(* IEC 61131-3 sources: SRCI_CLIENT_PLC/RobotLibrary/Library/POUs/_internal, 1 file *)

(* ---- ActiveCommandRegisterFB.st ---- *)
FUNCTION_BLOCK ActiveCommandRegisterFB EXTENDS RobotLibraryLogFB
// -------------------------------------------------------------------------
//  SRCI Robot Library
// -------------------------------------------------------------------------
//
//  Object:      ActiveCommandRegisterFB
//  Author:      Thorsten Brach
//  Date:        2024-06-01
//
//  Description:
//
//
//  Copyright:
//    (C) 2024 Thorsten Brach. All rights reserved
//             Licensed under the MIT License.
//
//  Disclaimer:
//    This project is provided without any guarantee and can be used for
//    private and commercial purposes. Any use is at the user’s
//    own risk and responsibility.
//
// -------------------------------------------------------------------------
VAR_INPUT
  /// Active Command Register
  Register            : ARRAY [1..RobotLibraryParameter.ACTIVE_CMD_REGISTER_ENTRIES_MAX] OF AxesGroupAcyclicAcrEntry;
  /// System Time
  SystemTime          : SystemTime;
  /// usable size of the arc register
  RegisterSize        : DINT := RobotLibraryParameter.ACTIVE_CMD_REGISTER_ENTRIES_MAX;
END_VAR

VAR_OUTPUT
  /// Execution Order List
  ExecutionOrderList    : ARRAY [1..RobotLibraryParameter.ACTIVE_CMD_REGISTER_ENTRIES_MAX] OF DINT;
  /// Current amount of used registers
  CurrentAcrUsageCount  : DINT;
  /// Current percent of used registers
  CurrentAcrUsagePercent : REAL;
END_VAR

VAR
  /// temporarty Active Command Register
  TmpRegister                 : ARRAY [1..RobotLibraryParameter.ACTIVE_CMD_REGISTER_ENTRIES_MAX] OF AxesGroupAcyclicAcrEntry;
  /// last used unique ID
  LastUniqueID                : UINT;
  /// Warning for ACR usage at 80%
  WarningAcrUsage             : R_TRIG;
END_VAR

VAR CONSTANT
  /// Active command
  ACTIVE_CMD           : UDINT := 1;
  /// Buffered command
  BUFFER_CMD           : UDINT := 2;
  /// Empty ACR entry
  EMPTY_ACR_ENTRY      : AxesGroupAcyclicAcrEntry := (State := ActiveCommandRegisterState.IS_FREE);
  /// Empty command entry
  EMPTY_CMD_ENTRY      : AxesGroupAcyclicAcrEntryCmdBuffer := (State := BufferStateCmd.EMPTY);
  /// constant for byte index of priority in payload
  PRIORITY_IDX         : BYTE := 3;
  /// bitmask to mask the priority out of the halfbyte
  PRIORITY_BIT_MASK    : BYTE := 2#000_1111;
END_VAR

  ManageRegister();

  UpdateExecutionOrderList();

END_FUNCTION_BLOCK

METHOD PUBLIC AddCmd : UDINT
VAR_INPUT
  /// Pointer to the corresponding command-FB to enable a callback mechanism
  pCommandFB        : POINTER TO RobotLibraryBaseFB;
END_VAR

VAR
  /// internal index for loops
 _regIdx            : DINT;
  /// internal command type
 _cmdType           : CmdType;
  /// log message
 _messageLog        : AlarmMessage;
  /// flag for free register found
 _freeRegisterFound : BOOL;
  /// internal Acr error
 _errorAcrEntry     : WORD := RobotLibraryErrorIdEnum.ERR_NO_FREE_ACR_ENTRY;
END_VAR

  // ST-FIX F48: a command with a parameter error of the block is not added
  IF ( pCommandFB <> 0 )
  THEN
    IF (( pCommandFB^.ErrorID = RobotLibraryErrorIdEnum.ERR_INVALID_PARAM_EXECUTION_MODE ) OR
        ( pCommandFB^.ErrorID = RobotLibraryErrorIdEnum.ERR_PROCESSINGMODE_NOT_DEFINED   ))
    THEN
      AddCmd := 0;
      RETURN;
    END_IF
  END_IF

  // calculate the used length of the ACR
  FOR _regIdx := 1 TO RegisterSize
  DO
    IF ( Register[_regIdx].State = ActiveCommandRegisterState.IS_FREE )
    THEN
      Register[_regIdx].State      := ActiveCommandRegisterState.IS_PROCESSING;
      Register[_regIdx].UniqueID   := DINT_TO_UINT(_regIdx);
      Register[_regIdx].pCommandFB := pCommandFB;

      // check pointer to command FB
      IF ( Register[_regIdx].pCommandFB <> RobotLibraryConstants.NULL_POINTER )
      THEN
        Register[_regIdx].Command[RobotLibraryConstants.ACTIVE_CMD].Timestamp  := SystemTime;

        Register[_regIdx].Command[RobotLibraryConstants.ACTIVE_CMD].Payload    := pCommandFB^.CommandData.Payload;
        Register[_regIdx].Command[RobotLibraryConstants.ACTIVE_CMD].PayloadLen := pCommandFB^.CommandData.PayloadLen;
        Register[_regIdx].Command[RobotLibraryConstants.ACTIVE_CMD].PayLoadPtr := 0;
        Register[_regIdx].Command[RobotLibraryConstants.ACTIVE_CMD].State      := BufferStateCmd.CREATED;
      END_IF

      // set flag for free register found
     _freeRegisterFound := TRUE;

      // Increment Current used register counter
      CurrentAcrUsageCount := CurrentAcrUsageCount + 1;

      // return Unique ID
      AddCmd := Register[_regIdx].UniqueID;

      // Get CmdType from payload
      SysDepMemCpy( pDest := ADR(_cmdType), pSrc := ADR(pCommandFB^.CommandData.Payload), DataLen := SIZEOF(_cmdType));

      // Create log entry
      CreateLogMessagePara2 ( Timestamp   := SystemTime,
                              MessageType := MessageType.CMD,
                              Severity    := Severity.INFO,
                              MessageCode := 0,
                              MessageText := 'ACR-ID [{1}]: Added  Command-Payload of CmdType <{2}>',
                              Para1       :=  DINT_TO_STRING(_regIdx),
                              Para2       :=  CMD_TYPE_TO_STRING(SwapUint(_cmdType)));
      EXIT;
    END_IF
  END_FOR

  // Check a free register could be found ?
  IF ( NOT _freeRegisterFound )
  THEN
    // set error in Command FB
    IF ( pCommandFB <> RobotLibraryConstants.NULL_POINTER )
    THEN
      SysDepMemCpy( pDest   := ADR   ( pCommandFB^.ErrorID ),
                    pSrc    := ADR   ( _errorAcrEntry      ),
                    DataLen := SIZEOF( _errorAcrEntry      ));
    END_IF

    // Create log entry
    CreateLogMessagePara1 ( Timestamp   := SystemTime,
                            MessageType := MessageType.CMD,
                            Severity    := Severity.FATAL_ERROR,
                            MessageCode := 0,
                            MessageText := 'Not possible to add CMD <{1}> to ACR - NO FREE REGISTER FOUND ! -> STOPPING SRCI INTERFACE...',
                            Para1       :=  CMD_TYPE_TO_STRING(SwapUint(_cmdType)));
  END_IF

END_METHOD

METHOD AddRsp : UDINT
VAR_INPUT
  /// Response
  Rsp : TelegramRobToPlcFragment;
END_VAR
VAR
  /// internal index for loops
 _Idx             : DINT;
  /// internal registen index
 _regIdx          : DINT;
  /// internal command type
 _cmdType         : CmdType;
  /// internal FragmentAction
 _fragmentAction  :  FragmentAction;
  /// internal command message state
 _cmdMessageState : CmdMessageState;
  /// internal flag for CmdID found
 _found           : BOOL;
END_VAR

  FOR _regIdx := 1 TO RegisterSize
  DO
    IF ( Register[_regIdx].UniqueID = Rsp.Header.CmdID )
    THEN
      // CmdID was found in the ACR
     _found := TRUE;
      // convert to fragment action
     _fragmentAction := ByteToFragmentAction(Rsp.Header.FragmentAction);

      // delete response
      IF ( _fragmentAction.Clear )
      THEN
        SysDepMemSet( pDest := ADR(Register[_regIdx].Response[ACTIVE_CMD]), Value := 0, DataLen := SIZEOF(Register[_regIdx].Response[ACTIVE_CMD]));
      END_IF

      // add payload to response
      FOR _idx := Rsp.Header.PayloadPointer TO  Rsp.Header.PayloadPointer + Rsp.Header.PayloadLength -1
      DO
        Register[_regIdx].Response[ACTIVE_CMD].Timestamp     := SystemTime;
        Register[_regIdx].Response[ACTIVE_CMD].State         := BufferStateRsp.RECEIVING;
        Register[_regIdx].Response[ACTIVE_CMD].PayloadLen    := Register[_regIdx].Response[ACTIVE_CMD].PayloadLen + 1;
        Register[_regIdx].Response[ACTIVE_CMD].Payload[_idx] := Rsp.Command.Payload[_idx];
      END_FOR

      // Get current message state
     _cmdMessageState := GetHalfeByteLo    (Value  := Register[_regIdx].Response[ACTIVE_CMD].Payload[0]);
      // Get command type from payload
     _cmdType         := CombineBytesToUint(HiByte := Register[_regIdx].Command [ACTIVE_CMD].Payload[0],
                                            LoByte := Register[_regIdx].Command [ACTIVE_CMD].Payload[1]);

      // Create log entry
      CreateLogMessagePara3 ( Timestamp   := SystemTime,
                              MessageType := MessageType.CMD,
                              Severity    := Severity.INFO,
                              MessageCode := 0,
                              MessageText := 'ACR-ID [{1}]: Added Response-Payload of CmdType <{2}> with State = {3}',
                              Para1       :=  DINT_TO_STRING(_regIdx),
                              Para2       :=  CMD_TYPE_TO_STRING(_cmdType),
                              Para3       :=  CMD_MESSAGE_STATE_TO_STRING(_cmdMessageState));

      IF ( _fragmentAction.Complete )
      THEN
        // set response state
        Register[_regIdx].Response[ACTIVE_CMD].State := BufferStateRsp.RECEIVED;

        // Check current message state and tag the register state as IS_FINAL, if needed
        IF ( _cmdMessageState >= CmdMessageState.DONE)
        THEN
          Register[_regIdx].State := ActiveCommandRegisterState.IS_FINAL;

          // get command type from payload
         _cmdType := CombineBytesToUint(HiByte := Register[_regIdx].Command[ACTIVE_CMD].Payload[0],
                                        LoByte := Register[_regIdx].Command[ACTIVE_CMD].Payload[1]);

          // Create log entry
          CreateLogMessagePara3( Timestamp   := SystemTime,
                                 MessageType := MessageType.CMD,
                                 Severity    := Severity.INFO,
                                 MessageCode := 0,
                                 MessageText := 'ACR-ID [{1}]: Detected Response-Payload of CmdType <{2}> has reached final state <{3}>',
                                 Para1       :=  DINT_TO_STRING(_regIdx),
                                 Para2       :=  CMD_TYPE_TO_STRING(_cmdType),
                                 Para3       :=  CMD_MESSAGE_STATE_TO_STRING(_cmdMessageState));

          // Exit the loop
        END_IF
      END_IF

      // Check Response received complete ?
      IF ( Register[_regIdx].Response[ACTIVE_CMD].State = BufferStateRsp.RECEIVED)
      THEN
        // update state
        Register[_regIdx].Response[ACTIVE_CMD].State := BufferStateRsp.PROCESSED;
        // callback CommandFB
        Register[_regIdx].pCommandFB^.CallBack(RspData := Register[_regIdx].Response[ACTIVE_CMD],TimeStamp := SystemTime);
      END_IF

      EXIT;
    END_IF
  END_FOR

  // Check CmdID was found in the ACR ?
  IF ( NOT _found )
  THEN
    // Create log entry
    CreateLogMessagePara2 ( Timestamp   := SystemTime,
                            MessageType := MessageType.CMD,
                            Severity    := Severity.WARNING,
                            MessageCode := 0,
                            MessageText := 'ACR-ID [?]: Response-Payload of CmdID <{1}> with State = {2} received, but no matching ACR entry found',
                            Para1       :=  UINT_TO_STRING(Rsp.Header.CmdID),
                            Para2       :=  CMD_MESSAGE_STATE_TO_STRING(_cmdMessageState));
  END_IF

END_METHOD

METHOD FB_init : BOOL
VAR_INPUT
  bInitRetains : BOOL; // if TRUE, the retain variables are initialized (warm start / cold start)
  bInCopyCode : BOOL;  // if TRUE, the instance afterwards gets moved into the copy code (online change)
END_VAR

  MyType := 'ActiveCommandRegisterFB';

END_METHOD

METHOD PRIVATE ManageRegister
VAR
  /// internal index
 _regIdx          : DINT;
  /// internal command type
 _cmdType         : CmdType;
  /// internal command message state
 _cmdMessageState : CmdMessageState;
END_VAR

  FOR _regIdx := 1 TO RegisterSize
  DO
    // Check pointer to command FB is valid ?
    IF ( Register[_regIdx].pCommandFB <> RobotLibraryConstants.NULL_POINTER)
    THEN

      // Check apply Cmd parameter update ?
      IF (( Register[_regIdx].Command[ACTIVE_CMD].State = BufferStateCmd.PROCESSED        ) AND
          ( Register[_regIdx].Command[BUFFER_CMD].State = BufferStateCmd.UPDATE_AVAILABLE ))
      THEN
        Register[_regIdx].Command[ACTIVE_CMD] := Register[_regIdx].Command[BUFFER_CMD];
        Register[_regIdx].Command[BUFFER_CMD] := EMPTY_CMD_ENTRY;

        // get command type from payload
       _cmdType := CombineBytesToUint(HiByte := Register[_regIdx].Command[ACTIVE_CMD].Payload[0],
                                      LoByte := Register[_regIdx].Command[ACTIVE_CMD].Payload[1]);

        // Create log entry
        CreateLogMessagePara2 ( Timestamp   := SystemTime,
                                MessageType := MessageType.CMD,
                                Severity    := Severity.INFO,
                                MessageCode := 0,
                                MessageText := 'ACR-ID [{1}]: Moved BUFFER_CMD to ACTIVE_CMD, CmdType <{2}>',
                                Para1       :=  DINT_TO_STRING(_regIdx),
                                Para2       :=  CMD_TYPE_TO_STRING(_cmdType));

      END_IF

      (*
      // Check Response received ?
      IF ( Register[_regIdx].Response[ACTIVE_CMD].State = BufferStateRsp.RECEIVED)
      THEN
        // update state
        Register[_regIdx].Response[ACTIVE_CMD].State := BufferStateRsp.PROCESSED;
        // callback CommandFB
        Register[_regIdx].pCommandFB^.CallBack(RspData := Register[_regIdx].Response[ACTIVE_CMD],TimeStamp := SystemTime);
      END_IF
      *)

      // delete entries with State.IS_Final
      IF ( Register[_regIdx].State = ActiveCommandRegisterState.IS_FINAL )
      THEN
        // get command type from payload
       _cmdType := CombineBytesToUint(HiByte := Register[_regIdx].Command[ACTIVE_CMD].Payload[0],
                                      LoByte := Register[_regIdx].Command[ACTIVE_CMD].Payload[1]);

        // Get current message state
       _cmdMessageState := GetHalfeByteLo(Value := Register[_regIdx].Response[ACTIVE_CMD].Payload[0]);

        // Create log entry
        CreateLogMessagePara3( Timestamp   := SystemTime,
                               MessageType := MessageType.CMD,
                               Severity    := Severity.INFO,
                               MessageCode := 0,
                               MessageText := 'ACR-ID [{1}]: Deleted ACR-Entry of CmdType <{2}> with State = {3}, because of Final-State was reached',
                               Para1       :=  DINT_TO_STRING(_regIdx),
                               Para2       :=  CMD_TYPE_TO_STRING(_cmdType),
                               Para3       :=  CMD_MESSAGE_STATE_TO_STRING(_cmdMessageState));

        // delete register entry
        Register[_regIdx] := EMPTY_ACR_ENTRY;

        // decrement current used register counter
        CurrentAcrUsageCount := CurrentAcrUsageCount - 1;
      END_IF
    END_IF
  END_FOR

  // Calculate percent of register usage
  IF ( CurrentAcrUsageCount > 0)
  THEN
    CurrentAcrUsagePercent :=  (DINT_TO_REAL(CurrentAcrUsageCount) / DINT_TO_REAL(RegisterSize)) * 100.0;
  ELSE
    CurrentAcrUsagePercent := 0.0;
  END_IF

  // build rising edge for arc usage over 80%
  WarningAcrUsage( CLK := CurrentAcrUsagePercent > RobotLibraryParameter.ACR_USAGE_WARNING_LIMIT );

  IF ( WarningAcrUsage.Q )
  THEN
    // Create log entry
    CreateLogMessagePara4( Timestamp   := SystemTime,
                           MessageType := MessageType.CMD,
                           Severity    := Severity.WARNING,
                           MessageCode := 0,
                           MessageText := 'ACR Register usage has reached the warning limit ({1}): {2}/{3} = {4}%',
                           Para1       :=  REAL_TO_STRING(RobotLibraryParameter.ACR_USAGE_WARNING_LIMIT),
                           Para2       :=  DINT_TO_STRING(CurrentAcrUsageCount),
                           Para3       :=  DINT_TO_STRING(RegisterSize),
                           Para4       :=  REAL_TO_STRING(CurrentAcrUsagePercent));
  END_IF

END_METHOD

PROPERTY PUBLIC NotifyParameterChanged : UDINT

SET
VAR
  /// internal register index
 _regIdx  : DINT;
  /// internal command type
 _cmdType : CmdType;
END_VAR

  FOR _regIdx := 1 TO RobotLibraryParameter.ACTIVE_CMD_REGISTER_ENTRIES_MAX
  DO
    // check unique ID found ?
    IF ( Register[_regIdx].UniqueID = NotifyParameterChanged )
    THEN
      // ST-FIX F114: a parameter change before the command is sent (state CREATED) must not turn the new
      // command into a parameter update (it was never sent): the command keeps the parameters of the rising edge
      IF ( Register[_regIdx].Command[ACTIVE_CMD].State = BufferStateCmd.CREATED )
      THEN
        // Create log entry
        CreateLogMessagePara1 ( Timestamp   := SystemTime,
                                MessageType := MessageType.CMD,
                                Severity    := Severity.INFO,
                                MessageCode := 0,
                                MessageText := 'ACR-ID [{1}]: Cmd-Parameter changed before the command was sent -> ignored',
                                Para1       :=  DINT_TO_STRING(_regIdx));
      ELSIF (( Register[_regIdx].Command[ACTIVE_CMD].State <> BufferStateCmd.SENDING   ) AND
             ( Register[_regIdx].Command[ACTIVE_CMD].State <> BufferStateCmd.PROCESSED ))
      THEN
        // Check pointer is valid ?
        IF ( Register[_regIdx].pCommandFB <> RobotLibraryConstants.NULL_POINTER )
        THEN
          // add to send register
          Register[_regIdx].Command[ACTIVE_CMD].Timestamp  := SystemTime;
          Register[_regIdx].Command[ACTIVE_CMD].State      := BufferStateCmd.UPDATE_AVAILABLE;
          Register[_regIdx].Command[ACTIVE_CMD].Payload    := Register[_regIdx].pCommandFB^.CommandData.Payload;
          Register[_regIdx].Command[ACTIVE_CMD].PayloadLen := Register[_regIdx].pCommandFB^.CommandData.PayloadLen;

          // get command type from payload
         _cmdType := CombineBytesToUint(HiByte := Register[_regIdx].pCommandFB^.CommandData.Payload[0],
                                        LoByte := Register[_regIdx].pCommandFB^.CommandData.Payload[1]);

          // Create log entry
          CreateLogMessagePara2 ( Timestamp   := SystemTime,
                                  MessageType := MessageType.CMD,
                                  Severity    := Severity.INFO,
                                  MessageCode := 0,
                                  MessageText := 'ACR-ID [{1}]: Updated Cmd-Parameter of CmdType <{2}> -> written to ACTIVE_CMD Index',
                                  Para1       :=  DINT_TO_STRING(_regIdx),
                                  Para2       :=  CMD_TYPE_TO_STRING(_cmdType));
        END_IF
      ELSE
        // Check pointer is valid ?
        IF ( Register[_regIdx].pCommandFB <> RobotLibraryConstants.NULL_POINTER )
        THEN
          // add to buffer register
          Register[_regIdx].Command[BUFFER_CMD].Timestamp  := SystemTime;
          Register[_regIdx].Command[BUFFER_CMD].State      := BufferStateCmd.UPDATE_AVAILABLE;
          Register[_regIdx].Command[BUFFER_CMD].Payload    := Register[_regIdx].pCommandFB^.CommandData.Payload;
          Register[_regIdx].Command[BUFFER_CMD].PayloadLen := Register[_regIdx].pCommandFB^.CommandData.PayloadLen;

          // get command type from payload
         _cmdType := CombineBytesToUint(HiByte := Register[_regIdx].pCommandFB^.CommandData.Payload[0],
                                        LoByte := Register[_regIdx].pCommandFB^.CommandData.Payload[1]);

          // Create log entry
          CreateLogMessagePara2 ( Timestamp   := SystemTime,
                                  MessageType := MessageType.CMD,
                                  Severity    := Severity.INFO,
                                  MessageCode := 0,
                                  MessageText := 'ACR-ID [{1}]: Updated Cmd-Parameter of CmdType <{2}> -> written to BUFFER_CMD Index',
                                  Para1       :=  DINT_TO_STRING(_regIdx),
                                  Para2       :=  CMD_TYPE_TO_STRING(_cmdType));
        END_IF
      END_IF

    END_IF
  END_FOR

END_SET

METHOD PUBLIC OnOnlineChange : DINT
VAR_INPUT
  /// unique ID
  UniqueID     : UDINT;
  /// Pointer to the corresponding command-FB to enable a callback mechanism
  pCommandFB   : POINTER TO RobotLibraryBaseFB;
END_VAR

VAR
  /// internal index for loops
 _regIdx : DINT;
END_VAR

  OnOnlineChange := -1;

  // Check command FB pointer is valid ?
  IF ( pCommandFB <> RobotLibraryConstants.NULL_POINTER)
  THEN
    FOR _regIdx := 1 TO RegisterSize
    DO
      // check unique ID found ?
      IF ( Register[_regIdx].UniqueID = UniqueID )
      THEN
        // update pointer to command FB
        Register[_regIdx].pCommandFB := pCommandFB;
        // Return result OK
        OnOnlineChange := RobotLibraryConstants.OK;
        EXIT;
      END_IF
    END_FOR
  END_IF

END_METHOD

METHOD PUBLIC RemoveCmd : DINT
VAR_INPUT
 /// unique ID
 UniqueID : UDINT;
END_VAR

VAR
  /// internal index
 _regIdx : DINT;
  /// internal command type
 _cmdType : CmdType;
END_VAR

  RemoveCmd := RobotLibraryConstants.HAS_ERROR;

  IF (UniqueID = 0)
  THEN
    UniqueID := UniqueID;
  END_IF

  FOR _regIdx := 1 TO RegisterSize
  DO
    // check unique ID found and not yet sended ?
    IF (( Register[_regIdx].UniqueID                  = UniqueID                        ) AND
        ( Register[_regIdx].Command[ACTIVE_CMD].State < BufferStateCmd.UPDATE_AVAILABLE ))
    THEN
      // Get CmdType from payload
      SysDepMemCpy( pDest := ADR(_cmdType), pSrc := ADR(Register[_regIdx].Command[ACTIVE_CMD].Payload), DataLen := SIZEOF(_cmdType));
      // delete register entry
      SysDepMemSet(pDest := ADR(Register[_regIdx]), Value := 0 , DataLen := SIZEOF(Register[_regIdx]));
      // decrement current used register counter
      CurrentAcrUsageCount := CurrentAcrUsageCount - 1;
      // Command successfull removed
      RemoveCmd := RobotLibraryConstants.OK;

      // Create log entry
      CreateLogMessagePara2 (  Timestamp   := SystemTime,
                               MessageType := MessageType.CMD,
                               Severity    := Severity.INFO,
                               MessageCode := 0,
                               MessageText := 'ACR-ID [{1}]: Removed CmdType <{2}>',
                               Para1       :=  DINT_TO_STRING(_regIdx),
                               Para2       :=  CMD_TYPE_TO_STRING(SwapUint(_cmdType)));
      EXIT;
    END_IF
  END_FOR

END_METHOD

METHOD PUBLIC Reset

  SysDepMemSet( ADR(Register), 0, SIZEOF(Register));

  CurrentAcrUsageCount   := 0;
  CurrentAcrUsagePercent := 0.0;

  // Create log entry
  CreateLogMessagePara1 ( Timestamp   := SystemTime,
                          MessageType := MessageType.CMD,
                          Severity    := Severity.INFO,
                          MessageCode := 0,
                          MessageText := 'ACR Registers has been reset and all entries deleted by Reset method call',
                          Para1       :=  '');

END_METHOD

METHOD PRIVATE UpdateExecutionOrderList
VAR
  /// temporary Active Command Register entry
  TmpRegisterEntry : AxesGroupAcyclicAcrEntry;
  /// temporary index
  TmpIndex         : DINT;
  /// internal index
  i                : DINT;
  /// internal index
  j                : DINT;
END_VAR

  // Reset temporary register
  SysDepMemSet(pDest := ADR(TmpRegister)       , Value := 0, DataLen := SIZEOF(TmpRegister));
  // Reset Execution Order List
  SysDepMemSet(pDest := ADR(ExecutionOrderList), Value := 0, DataLen := SIZEOF(ExecutionOrderList));
  // pre-set temporary register index
  j := 1;

  FOR i := 1 TO RegisterSize
  DO
    // add only entries which are not in status free and where datas must be processed
    IF (( Register[i].State                      > ActiveCommandRegisterState.IS_FREE ) AND
        ( Register[i].Command[ACTIVE_CMD].State <> BufferStateCmd.EMPTY               ) AND
        ( Register[i].Command[ACTIVE_CMD].State <> BufferStateCmd.PROCESSED           ))
    THEN
      // copy register entry
      TmpRegister[j] := Register[i];
      // store index of the entry from the ACR
      ExecutionOrderList[j] := i;
      // inc temporar register index
      j := j + 1;
    END_IF
  END_FOR

  // Bubble Sort to sort the priorities from the active command register
  FOR i := 1 TO RegisterSize
  DO
    FOR j := 1 TO RegisterSize - 1
    DO
      // check list entry is not empty ?
      IF (( TmpRegister[i  ].State = ActiveCommandRegisterState.IS_FREE ) OR
          ( TmpRegister[j+1].State = ActiveCommandRegisterState.IS_FREE ))
      THEN
        EXIT;
      END_IF

      IF (( TmpRegister[j].Command[ACTIVE_CMD].Payload[PRIORITY_IDX] AND PRIORITY_BIT_MASK ) > ( TmpRegister[j+1].Command[ACTIVE_CMD].Payload[PRIORITY_IDX] AND PRIORITY_BIT_MASK ))
      THEN
        // swap position of register entry
        TmpRegisterEntry := TmpRegister[j];
        TmpRegister[j]   := TmpRegister[j+1];
        TmpRegister[j+1] := TmpRegisterEntry;

        // swap position of index in the Execution Order List
        TmpIndex                := ExecutionOrderList[j];
        ExecutionOrderList[j]   := ExecutionOrderList[j+1];
        ExecutionOrderList[j+1] := TmpIndex;
      END_IF
    END_FOR
  END_FOR

  // Bubble Sort to sort the Timestamp from the pre-sorted active command register
  FOR i := 1 TO RegisterSize
  DO
    FOR j := 1 TO RegisterSize - 1
    DO
      // check list entry is not empty ?
      IF (( TmpRegister[i  ].State = ActiveCommandRegisterState.IS_FREE ) OR
          ( TmpRegister[j+1].State = ActiveCommandRegisterState.IS_FREE ))
      THEN
        EXIT;
      END_IF

         // Priority is higher
      IF (( TmpRegister[j].Command[ACTIVE_CMD].Payload[PRIORITY_IDX] AND PRIORITY_BIT_MASK ) >= ( TmpRegister[j+1].Command[ACTIVE_CMD].Payload[PRIORITY_IDX] AND PRIORITY_BIT_MASK )) AND
         // Date is greater
         (( TmpRegister[j].Command[ACTIVE_CMD].Timestamp.SystemDate                          >    TmpRegister[j+1].Command[ACTIVE_CMD].Timestamp.SystemDate                         ) OR
         // Date is the same, but Time is greater
         (( TmpRegister[j].Command[ACTIVE_CMD].Timestamp.SystemDate                          =    TmpRegister[j+1].Command[ACTIVE_CMD].Timestamp.SystemDate                         ) AND
          ( TmpRegister[j].Command[ACTIVE_CMD].Timestamp.SystemTime                          >    TmpRegister[j+1].Command[ACTIVE_CMD].Timestamp.SystemTime                         )))
      THEN
        // swap position of register entry
        TmpRegisterEntry := TmpRegister[j];
        TmpRegister[j]   := TmpRegister[j+1];
        TmpRegister[j+1] := TmpRegisterEntry;

        // swap position of index in the Execution Order List
        TmpIndex                := ExecutionOrderList[j];
        ExecutionOrderList[j]   := ExecutionOrderList[j+1];
        ExecutionOrderList[j+1] := TmpIndex;
      END_IF
    END_FOR
  END_FOR

END_METHOD
